(* IEC 61131-3 sources: codesys-framework/txt/application/WeVe Core (library)/70 Logger/I_Logger, 2 files *)

(* ---- LogEvent.method.st ---- *)
// Een event loggen. Wordt aangeroepen door FB_Event.
//   scEvent   : ID, level en bron (nSubMachine, nSubMachineId)
//   scPayload : de losse payloadvelden, voor gestructureerde loggers (Hyperion)
//   sMessage  : de volledige tekst, door het event opgebouwd
// TRUE = opgenomen in de buffer, FALSE = buffer vol (de logger telt de overflow).
METHOD LogEvent : BOOL
VAR_INPUT
	scEvent 		: SC_Event;
	scPayload 		: SC_EventPayload;
	sMessage 		: STRING(GVL_Logger.cMaxMessageLength);
END_VAR

(* ---- LogMessage.method.st ---- *)
// Vrije tekst loggen, bv. om te debuggen.
// TRUE = opgenomen in de buffer, FALSE = buffer vol (de logger telt de overflow).
METHOD LogMessage : BOOL
VAR_INPUT
	eLevel 			: E_EventLevels;
	sMessage 		: STRING(GVL_Logger.cMaxMessageLength);
END_VAR
